// TIA Portal V20 export
// export: Created 2026-10-12T18:08:14.8654693Z, ExportSetting WithDefaults, DisplayName Totally Integrated Automation Portal, DisplayVersion V20 Update 6, DisplayName TIA Portal Openness, DisplayVersion V20 Update 6, DisplayName TIA Portal Version Control Interface, DisplayVersion V20 Update 6, DisplayName SINAMICS Startdrive Advanced, DisplayVersion V20 SP1 Update 2, DisplayName SINAMICS Startdrive G110M, G120, G120C, G120D, G120P, G115D, DisplayVersion V20 SP1 Update 2, DisplayName SINAMICS Startdrive G130, G150, S120, S150, SINAMICS MV, G220, S200, S210, DisplayVersion V20 SP1 Update 2, DisplayName STEP 7 Professional, DisplayVersion V20 Update 6, DisplayName STEP 7 Safety, DisplayVersion V20 Update 2, DisplayName WinCC Basic/Comfort/Advanced, DisplayVersion V20 Update 6, DisplayName WinCC Professional, DisplayVersion V20 Update 6, DisplayName WinCC Unified, DisplayVersion V20 Update 6
FUNCTION_BLOCK "FB_Nachspeisung"   // FB2, SCL
{ S7_Optimized_Access := 'TRUE' }
VERSION : 0.1
// stored: AutoNumber true, IsIECCheckEnabled false, IsRetainMemResEnabled false, MemoryReserve 100, SetENOAutomatically false, UDAEnableTagReadback false
   VAR_INPUT
      Niveau_Bad_25_Roh : Bool;   // Sonde Bad 25, TRUE = Niveau OK (unverzoegert)
      Niveau_Bad_26_OK : Bool;   // Sonde Bad 26, TRUE = Niveau OK (Trockenlaufschutz)
      Motorschutz_OK : Bool;   // Motorschutz 275aQ1 und Wartungsschalter
      Not_Halt_Aktiv : Bool;
      Nachlaufzeit : Time;   // Nachlauf nach Niveau OK, aus DB_IPC_to_CPU
   END_VAR
   VAR_OUTPUT
      Pumpe_Ein : Bool;   // Ansteuerung 275aK8
      Niveau_Bad_25_OK : Bool;   // Niveau Bad 25 fuer die Badlogik, Fehler erst nach 30 s
      Zeitueberwachung_Stoerung : Bool;   // 5 min gepumpt, Niveau Bad 25 immer noch nicht OK
   END_VAR
   VAR
      Timer_Niveau_25 { S7_SetPoint := 'True'} : TON_TIME;
      Timer_Anforderung { S7_SetPoint := 'True'} : TON_TIME;
      Timer_Quelle { S7_SetPoint := 'True'} : TON_TIME;
      Timer_Nachlauf { S7_SetPoint := 'True'} : TON_TIME;
      Timer_Laufzeit { S7_SetPoint := 'True'} : TON_TIME;
      Anforderung_Aktiv : Bool;
      Stoerung : Bool;
   END_VAR
   VAR_TEMP
      nachlauf : Time;
      freigabe : Bool;
   END_VAR
BEGIN

       //== 1) Niveau Bad 25 fuer die Badlogik: Fehler erst wenn 30 s nicht OK ==
       #Timer_Niveau_25(IN := NOT #Niveau_Bad_25_Roh, PT := T#30s);
       #Niveau_Bad_25_OK := NOT #Timer_Niveau_25.Q;

       //== 2) Nachlaufzeit (negative Werte wie 0 behandeln) ==
       IF #Nachlaufzeit < T#0s THEN #nachlauf := T#0s; ELSE #nachlauf := #Nachlaufzeit; END_IF;

       //== 3) Freigabe: Niveau Bad 26 mind. 5 s OK (Abfall sofort = Trockenlaufschutz), Motorschutz, kein Not-Halt ==
       #Timer_Quelle(IN := #Niveau_Bad_26_OK, PT := T#5s);
       #freigabe := #Timer_Quelle.Q AND #Motorschutz_OK AND NOT #Not_Halt_Aktiv;

       //== 4) Anforderung: Niveau Bad 25 5 s nicht OK -> an; Niveau OK + Nachlaufzeit -> aus ==
       #Timer_Anforderung(IN := NOT #Niveau_Bad_25_Roh, PT := T#5s);
       IF #Anforderung_Aktiv THEN
           #Timer_Nachlauf(IN := #Niveau_Bad_25_Roh, PT := #nachlauf);
           IF #Timer_Nachlauf.Q THEN #Anforderung_Aktiv := FALSE; END_IF;
       ELSE
           #Timer_Nachlauf(IN := FALSE, PT := #nachlauf);
           IF #Timer_Anforderung.Q AND NOT #Stoerung THEN #Anforderung_Aktiv := TRUE; END_IF;
       END_IF;

       //== 5) Pumpe ==
       #Pumpe_Ein := #Anforderung_Aktiv AND #freigabe AND NOT #Stoerung;

       //== 6) Zeitueberwachung: 5 min gepumpt und Niveau Bad 25 immer noch nicht OK ==
       #Timer_Laufzeit(IN := #Pumpe_Ein AND NOT #Niveau_Bad_25_Roh, PT := T#5m);
       IF #Timer_Laufzeit.Q THEN
           #Stoerung := TRUE;
           #Anforderung_Aktiv := FALSE;
       END_IF;
       // automatische Quittierung: Niveau Bad 25 wieder OK
       IF #Stoerung AND #Niveau_Bad_25_Roh THEN
           #Stoerung := FALSE;
       END_IF;
       #Pumpe_Ein := #Pumpe_Ein AND NOT #Stoerung;

       #Zeitueberwachung_Stoerung := #Stoerung;
END_FUNCTION_BLOCK
